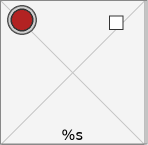
VISUALIZATION Vis_ES_PB  // 148x145
VAR_IN_OUT
	stPB: ST_ES_PB;

END_VAR
VAR_INPUT
	Lable: STRING;

END_VAR
    Image (0,0 145x145), "%s", text variable: Lable, image: ImagePool.EStop_OK2
        p84334746: stPB.stBitMap
    Checkbox (107,3 41x39), tooltip "ByPass", variable: stPB.ByPass, input disabled if: prg_User.actUser<4
    Lamp1 (5,3 34x34), tooltip "Memo PB State", variable: stPB.Memo, style: Lamp-Lamp1-Red
END_VISUALIZATION

(* stored: Version 1.1.0.1, ProductVersion 3.1.4024.13
   Visu Vis_ES_PB: Id {392dc3d7-debf-4965-9520-c9c46e3f1c39} *)
